(* IEC 61131-3 sources: stdmachine/plc/src/05_Sequencers, 11 files *)

(* ---- GVL_Active.st ---- *)
// Zone active du déploiement (docs/05 § 9 et § 10) : persistante, le PLC redémarre Stopped avec le dernier
// déploiement. À vérifier sur la cible : la taille (environ 1,5 Mo) des données persistantes.
{attribute 'qualified_only'}
VAR_GLOBAL PERSISTENT
    stMachine : ST_MachineData;
    aStation : ARRAY[1..GVL_Const.MAX_STATIONS] OF ST_StationData;
    aPressRecipe : ARRAY[1..GVL_Const.MAX_PRESS_RECIPES] OF ST_PressRecipe;
    bDeployed : BOOL;               // un déploiement a été activé
    nRetainId : ULINT;              // identifiant de la mémoire rémanente (docs/02 § 7.4), tiré au premier démarrage
END_VAR

(* ---- FB_GeneralSequencer.st ---- *)
// Séquenceur général (docs/05 § 5) : exécution du process général par mover, routage vers les stations des
// fonctions, files et priorités, préparation, fin d'opération (création et clôture des pièces, traces, qualité),
// table d'OF, fin des pièces en cours, variables de mover, mover à vider, mover hors service.
FUNCTION_BLOCK FB_GeneralSequencer
VAR_INPUT
    bDrain : BOOL;                  // fin des pièces en cours (docs/05 § 5.7), posé et levé par FB_Machine
END_VAR
VAR_OUTPUT
    bStopRequest : BOOL;            // impulsion : arrêt automatique demandé à la machine
    nStopReason : UINT;             // 1 OF terminé, 2 machine vidée, 3 arrêt qualité
    bMachineFault : BOOL;           // mover en défaut, alarme de process « défaut machine »
    nFaultCode : UINT;
END_VAR
VAR
    _refMachine : REFERENCE TO ST_MachineData;
    _refMgr : REFERENCE TO FB_MoverManager;
    _refQuality : REFERENCE TO FB_QualityMonitor;
    _refAlarms : REFERENCE TO FB_AlarmManager;
    _refTraces : REFERENCE TO FB_TraceBuffer;
    aStation : ARRAY[1..GVL_Const.MAX_STATIONS] OF POINTER TO FB_Station;
    _aLastReceived : ARRAY[1..GVL_Const.MAX_STATIONS] OF LINT;
    _aNoStationMs : ARRAY[1..GVL_Const.MAX_MOVERS] OF LREAL;
    _bExecute : BOOL;
    _bOrderDonePending : BOOL;      // l'OF actif vient de passer Done : arrêt quand plus aucune pièce
    _aGroupUsed : ARRAY[1..GVL_Const.MAX_GROUPS] OF BOOL;     // fonctions visées par une Route du process général
END_VAR
VAR PERSISTENT
    aMover : ARRAY[1..GVL_Const.MAX_MOVERS] OF ST_MoverCtx;
    aOrder : ARRAY[1..GVL_Const.MAX_ORDERS] OF ST_OrderState;
    nActiveOrder : USINT;           // rang dans aOrder, 0 = aucun
    _nReqSeq : UDINT;
    _nPartCounter : UDINT;
END_VAR

// ================================================================== mise en place

METHOD Init
VAR_INPUT
    refMachine : REFERENCE TO ST_MachineData;
    refMgr : REFERENCE TO FB_MoverManager;
    refQuality : REFERENCE TO FB_QualityMonitor;
    refAlarms : REFERENCE TO FB_AlarmManager;
    refTraces : REFERENCE TO FB_TraceBuffer;
END_VAR
_refMachine REF= refMachine;
_refMgr REF= refMgr;
_refQuality REF= refQuality;
_refAlarms REF= refAlarms;
_refTraces REF= refTraces;
END_METHOD

METHOD SetStation
VAR_INPUT
    nStation : USINT;
    pStation : POINTER TO FB_Station;
END_VAR
IF nStation >= 1 AND nStation <= GVL_Const.MAX_STATIONS THEN aStation[nStation] := pStation; END_IF
END_METHOD

// Reset machine (docs/05 § 6.3) : chaque mover détecté reçoit sa position ; les contextes et les pièces sont gardés
METHOD OnReset
VAR
    i : USINT;
    nPos : INT;
    ipDrv : I_PlanarDriver;
END_VAR
ipDrv := _refMgr.Driver;
FOR i := 1 TO _refMachine.nMovers DO
    aMover[i].bAbsent := FALSE;
    IF ipDrv <> 0 THEN
        IF NOT ipDrv.MoverDetected(i) THEN
            aMover[i].bAbsent := aMover[i].bOutOfService;       // D85 : un mover hors service peut être absent
            IF aMover[i].bAbsent AND __ISVALIDREF(_refAlarms) THEN _refAlarms.RaiseEvent(0, 915, i, E_Severity.Info); END_IF
        END_IF
    END_IF
    nPos := _refMgr.PositionAt(i);
    _refMgr.FreeAll(i, nPos);
    IF nPos > 0 THEN _refMgr.Reserve(nPos, i); END_IF
    aMover[i].nPos := nPos;
    CASE aMover[i].eState OF
        E_MoverState.Routing, E_MoverState.Halted, E_MoverState.Unknown, E_MoverState.Error:
            aMover[i].eState := E_MoverState.Ready;             // la Route en cours est reprise au Start
        E_MoverState.Queued:
            aMover[i].eState := E_MoverState.Buffered;
        E_MoverState.AtStation:
            IF NOT aMover[i].bStationAborted THEN
                aMover[i].eState := E_MoverState.Ready;
                aMover[i].bRequestPosted := FALSE;
            END_IF
    END_CASE
    IF aMover[i].nTable = 0 THEN
        aMover[i].nTable := 1;
        aMover[i].nPC := _refMachine.aTable[1].nStart;
    END_IF
END_FOR
END_METHOD

// Nouveau déploiement (docs/05 § 10) : variables de mover reprises par identifiant et type ; movers remis à
// l'étape 1 si le process général a changé de taille
METHOD OnDeploy
VAR_INPUT
    bRestartMovers : BOOL;
END_VAR
VAR
    i : USINT;
    v : USINT;
    k : USINT;
    stOld : ST_MoverCtx;
    bFound : BOOL;
END_VAR
FOR i := 1 TO GVL_Const.MAX_MOVERS DO
    stOld := aMover[i];
    FOR v := 1 TO GVL_Const.MAX_MOVER_VARS DO
        aMover[i].aVar[v] := 0;
        MEMSET(ADR(aMover[i].aVarPos[v]), 0, SIZEOF(ST_Position));
        aMover[i].aVarId[v] := 0;
        IF v <= _refMachine.nMoverVar THEN
            aMover[i].aVarId[v] := _refMachine.aMoverVar[v].nId;
            aMover[i].aVar[v] := _refMachine.aMoverVar[v].fInit;
            aMover[i].aVarPos[v] := _refMachine.aMoverVar[v].stInitPos;
            bFound := FALSE;
            IF _refMachine.aMoverVar[v].eReset <> E_MoverVarReset.OnDeploy THEN
                FOR k := 1 TO GVL_Const.MAX_MOVER_VARS DO
                    IF NOT bFound AND stOld.aVarId[k] = _refMachine.aMoverVar[v].nId AND stOld.aVarId[k] <> 0 THEN
                        aMover[i].aVar[v] := stOld.aVar[k];
                        aMover[i].aVarPos[v] := stOld.aVarPos[k];
                        bFound := TRUE;
                    END_IF
                END_FOR
            END_IF
        END_IF
    END_FOR
    IF bRestartMovers OR i > _refMachine.nMovers THEN
        aMover[i].nTable := 1;
        aMover[i].nPC := _refMachine.aTable[1].nStart;
        aMover[i].nDepth := 0;
        aMover[i].eState := E_MoverState.Ready;
        aMover[i].nTargetGroup := 0;
        aMover[i].bRequestPosted := FALSE;
    END_IF
END_FOR
IF bRestartMovers AND __ISVALIDREF(_refAlarms) THEN _refAlarms.RaiseEvent(0, 916, _refMachine.nMovers, E_Severity.Info); END_IF
ScanGroups();
END_METHOD

// ================================================================== cycle

METHOD Cycle
VAR_INPUT
    eState : E_State;               // état de la machine
END_VAR
VAR
    n : USINT;
    i : USINT;
    nArr : INT;
    nOldest : USINT;
END_VAR
_bExecute := eState = E_State.Execute;
bStopRequest := FALSE;
// Ordre des n°, en commençant par le mover qui attend depuis le plus longtemps (pas de famine)
nOldest := 1;
FOR i := 1 TO _refMachine.nMovers DO
    IF (aMover[i].eState = E_MoverState.Buffered OR aMover[i].eState = E_MoverState.Queued)
       AND (NOT (aMover[nOldest].eState = E_MoverState.Buffered OR aMover[nOldest].eState = E_MoverState.Queued) OR aMover[i].tWaitStart < aMover[nOldest].tWaitStart) THEN
        nOldest := i;
    END_IF
END_FOR
FOR n := 1 TO _refMachine.nMovers DO
    i := ((nOldest - 1 + n - 1) MOD _refMachine.nMovers) + 1;
    // Arrivées et timeouts, dans tous les états
    nArr := _refMgr.Arrived(i);
    IF nArr > 0 THEN _Arrive(i, nArr); END_IF
    IF _refMgr.TimedOut(i) AND aMover[i].eState <> E_MoverState.Error THEN
        aMover[i].eState := E_MoverState.Error;
        bMachineFault := TRUE;
        nFaultCode := 914;
        IF __ISVALIDREF(_refAlarms) THEN _refAlarms.RaiseEvent(0, 914, i, E_Severity.MachineFault); END_IF
    END_IF
    // Réaction qualité « mover hors service » (docs/10 § 5.1)
    aMover[i].bQualityLock := _refQuality.aMoverOut[i];

    IF _bExecute THEN
        IF (aMover[i].bOutOfService OR aMover[i].bQualityLock) AND aMover[i].eState = E_MoverState.Ready AND _Empty(i) THEN
            _SendToPark(i, FALSE);
        ELSIF aMover[i].bOutOfService AND aMover[i].bImmediate AND aMover[i].eState = E_MoverState.Ready AND NOT _Empty(i) THEN
            _SendToPark(i, TRUE);
        END_IF
        CASE aMover[i].eState OF
            E_MoverState.Ready: _RunMover(i);
            E_MoverState.Buffered:
                IF aMover[i].nTargetGroup = 0 THEN aMover[i].eState := E_MoverState.Ready; ELSE _TryRoute(i); END_IF
            E_MoverState.Queued: _Queued(i);
            E_MoverState.AtStation: _AtStation(i);
            E_MoverState.Halted: _Resume(i);
            E_MoverState.OutOfService:
                IF NOT aMover[i].bOutOfService AND NOT aMover[i].bQualityLock THEN _Restart(i); END_IF
        END_CASE
    ELSE
        // Held, Stopping : plus de nouveau routage ; les opérations lancées se terminent (docs/05 § 5.3)
        IF aMover[i].eState = E_MoverState.AtStation THEN _AtStation(i);
        ELSIF aMover[i].eState = E_MoverState.Ready OR aMover[i].eState = E_MoverState.Buffered OR aMover[i].eState = E_MoverState.Queued THEN
            IF eState = E_State.Held OR eState = E_State.Stopping THEN aMover[i].eWait := E_WaitReason.Held; END_IF
        END_IF
    END_IF
END_FOR
_CheckOrders();
IF bDrain AND (_bExecute OR eState = E_State.Held) AND PartsInProcess() = 0 AND NOT EntryInProgress() THEN
    bStopRequest := TRUE;
    nStopReason := 2;                                   // machine vidée (docs/05 § 5.7)
END_IF
IF _refQuality.bMachineStop THEN
    bStopRequest := TRUE;
    nStopReason := 3;
END_IF
_Publish();
END_METHOD

// ================================================================== process général d'un mover (docs/05 § 5.3)

METHOD PRIVATE _RunMover
VAR_INPUT
    i : USINT;
END_VAR
VAR
    m : REFERENCE TO ST_MoverCtx;
    ins : REFERENCE TO ST_Instr;
    nGuard : INT;
    n : INT;
    eSev : E_Severity;
END_VAR
m REF= aMover[i];
FOR nGuard := 1 TO 64 DO
    IF m.nPC < 1 OR m.nPC > _refMachine.nInstrCount THEN
        m.nTable := 1;
        m.nPC := _refMachine.aTable[1].nStart;
        RETURN;
    END_IF
    ins REF= _refMachine.aInstr[m.nPC];
    CASE ins.eOp OF
        E_Op.Jump:
            m.nPC := DINT_TO_INT(ins.aArg[1]);
        E_Op.JumpIfFalse:
            _MarkVerdictTested(i, DINT_TO_INT(ins.aArg[1]));
            IF _EvalCond(i, DINT_TO_INT(ins.aArg[1])) THEN m.nPC := m.nPC + 1; ELSE m.nPC := DINT_TO_INT(ins.aArg[2]); END_IF
        E_Op.SetVar:
            _SetVar(i);
            m.nPC := m.nPC + 1;
        E_Op.ResetMoverVars:
            _ResetVars(i, DINT_TO_INT(ins.aArg[1]));
            m.nPC := m.nPC + 1;
        E_Op.LoopInit:
            n := LIMIT(1, DINT_TO_INT(ins.aArg[1]), 8);
            m.aHidden[n] := _Resolve(i, ins.aParam[1]);
            m.nPC := m.nPC + 1;
        E_Op.LoopNext:
            n := LIMIT(1, DINT_TO_INT(ins.aArg[1]), 8);
            m.aHidden[n] := m.aHidden[n] - 1;
            IF m.aHidden[n] > 0 THEN m.nPC := DINT_TO_INT(ins.aArg[2]); ELSE m.nPC := m.nPC + 1; END_IF
        E_Op.Call:
            IF m.nDepth >= GVL_Const.MAX_CALL_DEPTH THEN
                m.eState := E_MoverState.Error;
                bMachineFault := TRUE;
                nFaultCode := 904;
                IF __ISVALIDREF(_refAlarms) THEN _refAlarms.RaiseEvent(0, 904, i, E_Severity.MachineFault); END_IF
                RETURN;
            END_IF
            m.nDepth := m.nDepth + 1;
            m.aRetTable[m.nDepth] := m.nTable;
            m.aRetPC[m.nDepth] := m.nPC + 1;
            m.nTable := DINT_TO_INT(ins.aArg[1]);
            m.nPC := _refMachine.aTable[m.nTable].nStart;
        E_Op.Return:
            IF m.nDepth = 0 THEN
                m.nTable := 1;
                m.nPC := _refMachine.aTable[1].nStart;
                RETURN;
            END_IF
            m.nTable := m.aRetTable[m.nDepth];
            m.nPC := m.aRetPC[m.nDepth];
            m.nDepth := m.nDepth - 1;
        E_Op.Alarm:
            // aArg[2] : 1 avertissement, sinon défaut machine (pas de station au niveau machine)
            IF ins.aArg[2] = 1 THEN eSev := E_Severity.Warning; ELSE eSev := E_Severity.MachineFault; END_IF
            IF __ISVALIDREF(_refAlarms) THEN _refAlarms.RaiseEvent(0, DINT_TO_UINT(ins.aArg[3]), i, eSev); END_IF
            IF ins.aArg[2] >= 2 THEN
                m.eState := E_MoverState.Error;
                bMachineFault := TRUE;
                nFaultCode := DINT_TO_UINT(ins.aArg[3]);
                RETURN;
            END_IF
            m.nPC := m.nPC + 1;
        E_Op.WaitCond:
            IF NOT _EvalCond(i, DINT_TO_INT(ins.aArg[1])) THEN RETURN; END_IF
            m.nPC := m.nPC + 1;
        E_Op.End:
            IF NOT _Empty(i) AND __ISVALIDREF(_refAlarms) THEN _refAlarms.RaiseEvent(0, 910, i, E_Severity.Warning); END_IF
            m.nTable := 1;
            m.nDepth := 0;
            m.nPC := _refMachine.aTable[1].nStart;
            RETURN;                                     // un tour de process par cycle au plus
        E_Op.Route:
            _StartRoute(i);
            RETURN;
    ELSE
        m.nPC := m.nPC + 1;                             // Nop, StepBegin, StepEnd
    END_CASE
END_FOR
END_METHOD

// ================================================================== routage (docs/05 § 5.4)

METHOD PRIVATE _StartRoute
VAR_INPUT
    i : USINT;
END_VAR
VAR
    m : REFERENCE TO ST_MoverCtx;
    ins : REFERENCE TO ST_Instr;
    nGroup : USINT;
    k : USINT;
    s : USINT;
    bBad : BOOL;
    bHandled : BOOL;
END_VAR
m REF= aMover[i];
ins REF= _refMachine.aInstr[m.nPC];
nGroup := DINT_TO_USINT(ins.aArg[1]);
m.nTargetOp := DINT_TO_USINT(ins.aArg[2]);
m.nTargetSlot := DINT_TO_USINT(ins.aArg[3]);
// 1. Pièce mauvaise non traitée par le process : redirection vers la fonction de rebut
FOR s := 1 TO GVL_Const.MAX_SLOTS DO
    IF m.aSlot[s].bPresent THEN
        bBad := bBad OR m.aSlot[s].aData[1] = 2;
        bHandled := bHandled OR m.aSlot[s].bBadHandled;
    END_IF
END_FOR
IF _refMachine.nRejectGroup > 0 AND nGroup <> _refMachine.nRejectGroup AND bBad AND NOT bHandled
   AND nGroup >= 1 AND nGroup <= GVL_Const.MAX_GROUPS AND_THEN _refMachine.aGroup[nGroup].eRole <> E_GroupRole.Reject THEN
    nGroup := _refMachine.nRejectGroup;
    m.nTargetOp := 1;
    MEMSET(ADR(m.aOpParam), 0, SIZEOF(m.aOpParam));
ELSE
    FOR k := 1 TO GVL_Const.MAX_PARAMS DO m.aOpParam[k] := _Resolve(i, ins.aParam[k]); END_FOR
END_IF
m.nTargetGroup := nGroup;
m.nStation := 0;
_aNoStationMs[i] := 0;
_TryRoute(i);
END_METHOD

METHOD PRIVATE _TryRoute
VAR_INPUT
    i : USINT;
END_VAR
VAR
    m : REFERENCE TO ST_MoverCtx;
    g : REFERENCE TO ST_GroupCfg;
    s : USINT;
    nBest : USINT;
    nLoad : INT;
    nBestLoad : INT;
    nDest : INT;
    k : USINT;
    eWait : E_WaitReason;
END_VAR
m REF= aMover[i];
IF m.nTargetGroup < 1 OR m.nTargetGroup > GVL_Const.MAX_GROUPS THEN m.eState := E_MoverState.Ready; RETURN; END_IF
g REF= _refMachine.aGroup[m.nTargetGroup];
// Fonction d'entrée : pas de chargement sans OF actif, OF complet, arrêt qualité du chargement, fin des pièces
IF g.eRole = E_GroupRole.Entry THEN
    eWait := _LoadingLock();
    IF eWait <> E_WaitReason.None THEN _WaitInBuffer(i, eWait); RETURN; END_IF
END_IF
// Candidates : stations membres en Execute, sans défaut, sans arrêt qualité, en production
nBest := 0;
IF NOT m.bOutOfService AND NOT m.bQualityLock THEN
    FOR s := 1 TO GVL_Const.MAX_STATIONS DO
        IF (SHR(g.nStationMask, s - 1) AND 1) = 1 AND_THEN _Routable(s) THEN
            nLoad := _LoadOf(s);
            IF nBest = 0 OR nLoad < nBestLoad OR (nLoad = nBestLoad AND _aLastReceived[s] < _aLastReceived[nBest]) THEN
                nBest := s;
                nBestLoad := nLoad;
            END_IF
        END_IF
    END_FOR
END_IF
IF nBest = 0 THEN
    _aNoStationMs[i] := _aNoStationMs[i] + F_CycleMs();
    IF (g.eRole = E_GroupRole.Reject OR _refMachine.nRejectGroup = 0) AND _aNoStationMs[i] > UDINT_TO_LREAL(_refMachine.nNoStationMs) AND NOT _Empty(i) THEN
        _SendToPark(i, TRUE);                       // mover à vider (911)
        RETURN;
    END_IF
    _WaitInBuffer(i, E_WaitReason.NoStation);
    RETURN;
END_IF
_aNoStationMs[i] := 0;
// Destination : position de travail libre et sans file, sinon une place de file, sinon un tampon
nDest := 0;
// (une position déjà tenue par ce mover compte comme libre : reprise après Reset)
IF _refMachine.aStation[nBest].nWorkPos > 0 AND_THEN _FreeFor(_refMachine.aStation[nBest].nWorkPos, i) AND NOT _HasQueue(nBest) THEN
    nDest := _refMachine.aStation[nBest].nWorkPos;
ELSE
    FOR k := 1 TO GVL_Const.MAX_QUEUE DO
        IF nDest = 0 AND _refMachine.aStation[nBest].aQueuePos[k] > 0 AND_THEN _FreeFor(_refMachine.aStation[nBest].aQueuePos[k], i) THEN
            nDest := _refMachine.aStation[nBest].aQueuePos[k];
        END_IF
    END_FOR
END_IF
IF nDest = 0 THEN
    _WaitInBuffer(i, E_WaitReason.NoStation);
    RETURN;
END_IF
_aLastReceived[nBest] := F_NowUtc();
m.nStation := nBest;
m.eWait := E_WaitReason.None;
IF _refMgr.MoveTo(i, nDest) THEN
    m.nDest := nDest;
    m.nPos := 0;
    m.eState := E_MoverState.Routing;
    m.bRequestPosted := FALSE;
    // Préparation : la demande est posée dès la réservation de la position de travail (docs/05 § 4.1)
    IF nDest = _refMachine.aStation[nBest].nWorkPos THEN _PostIfPrepare(i); END_IF
END_IF
END_METHOD

METHOD PRIVATE _FreeFor : BOOL
VAR_INPUT
    nPos : INT;
    i : USINT;
END_VAR
_FreeFor := _refMgr.Owner(nPos) = 0 OR _refMgr.Owner(nPos) = i;
END_METHOD

METHOD PRIVATE _LoadingLock : E_WaitReason
_LoadingLock := E_WaitReason.None;
IF _refQuality.bLoadingLocked THEN _LoadingLock := E_WaitReason.QualityStop;
ELSIF bDrain THEN _LoadingLock := E_WaitReason.Drain;
ELSIF nActiveOrder = 0 THEN _LoadingLock := E_WaitReason.NoOrder;
ELSIF aOrder[nActiveOrder].nGood + aOrder[nActiveOrder].nInProcess >= aOrder[nActiveOrder].nQuantity THEN _LoadingLock := E_WaitReason.OrderComplete;
END_IF
END_METHOD

METHOD PRIVATE _Routable : BOOL
VAR_INPUT
    s : USINT;
END_VAR
IF aStation[s] = 0 THEN _Routable := FALSE; RETURN; END_IF
_Routable := aStation[s]^.State = E_State.Execute AND NOT aStation[s]^.OutOfProduction AND NOT aStation[s]^.QualityLock
             AND _refMachine.aStation[s].bUsed;
END_METHOD

METHOD PRIVATE _LoadOf : INT
VAR_INPUT
    s : USINT;
END_VAR
VAR
    i : USINT;
END_VAR
_LoadOf := 0;
FOR i := 1 TO _refMachine.nMovers DO
    IF aMover[i].nStation = s THEN _LoadOf := _LoadOf + 1; END_IF
END_FOR
END_METHOD

METHOD PRIVATE _HasQueue : BOOL
VAR_INPUT
    s : USINT;
END_VAR
VAR
    i : USINT;
END_VAR
_HasQueue := FALSE;
FOR i := 1 TO _refMachine.nMovers DO
    IF aMover[i].nStation = s AND aMover[i].eState = E_MoverState.Queued THEN _HasQueue := TRUE; END_IF
END_FOR
END_METHOD

METHOD PRIVATE _WaitInBuffer
VAR_INPUT
    i : USINT;
    eReason : E_WaitReason;
END_VAR
VAR
    m : REFERENCE TO ST_MoverCtx;
    nBuf : INT;
END_VAR
m REF= aMover[i];
IF m.eState <> E_MoverState.Buffered THEN m.tWaitStart := F_NowUtc(); END_IF
m.eWait := eReason;
m.nStation := 0;
// Déjà sur un tampon ou au parcage : il y reste
IF m.nPos > 0 AND_THEN (_refMachine.aPlanarPos[m.nPos].eKind = E_PlanarPosKind.Buffer OR _refMachine.aPlanarPos[m.nPos].eKind = E_PlanarPosKind.Park) THEN
    m.eState := E_MoverState.Buffered;
    RETURN;
END_IF
IF m.eState = E_MoverState.Routing THEN RETURN; END_IF
nBuf := _refMgr.NearestFree(i, E_PlanarPosKind.Buffer);
IF nBuf > 0 AND_THEN _refMgr.MoveTo(i, nBuf) THEN
    m.nDest := nBuf;
    m.nPos := 0;
    m.eState := E_MoverState.Routing;
ELSE
    m.eState := E_MoverState.Buffered;                      // aucun tampon libre : il reste où il est
END_IF
END_METHOD

METHOD PRIVATE _SendToPark
VAR_INPUT
    i : USINT;
    bToEmpty : BOOL;
END_VAR
VAR
    m : REFERENCE TO ST_MoverCtx;
    nPark : INT;
END_VAR
m REF= aMover[i];
m.nStation := 0;
m.bToEmptyPark := bToEmpty;
IF bToEmpty AND __ISVALIDREF(_refAlarms) THEN _refAlarms.Raise(0, 911, i, E_Severity.Warning); END_IF
nPark := _refMachine.nParkPos;
IF nPark = 0 OR m.nPos = nPark THEN
    m.eState := SEL(bToEmpty OR NOT _Empty(i), E_MoverState.OutOfService, E_MoverState.ToEmpty);
    RETURN;
END_IF
IF _refMgr.MoveTo(i, nPark) THEN
    m.nDest := nPark;
    m.nPos := 0;
    m.eState := E_MoverState.Routing;
END_IF
END_METHOD

METHOD PRIVATE _Arrive
VAR_INPUT
    i : USINT;
    nPos : INT;
END_VAR
VAR
    m : REFERENCE TO ST_MoverCtx;
END_VAR
m REF= aMover[i];
m.nPos := nPos;
m.nDest := 0;
CASE _refMachine.aPlanarPos[nPos].eKind OF
    E_PlanarPosKind.Work:
        m.eState := E_MoverState.AtStation;
        IF m.bRequestPosted AND m.nStation >= 1 AND_THEN aStation[m.nStation] <> 0 THEN aStation[m.nStation]^.MoverArrived(m.nReqId); END_IF
    E_PlanarPosKind.Queue:
        // En Held et Stopping, le mover arrivé passe Halted (docs/05 § 5.3)
        IF _bExecute THEN m.eState := E_MoverState.Queued; ELSE m.eState := E_MoverState.Halted; END_IF
    E_PlanarPosKind.Buffer:
        IF _bExecute THEN m.eState := E_MoverState.Buffered; ELSE m.eState := E_MoverState.Halted; END_IF
    E_PlanarPosKind.Park:
        IF m.bToEmptyPark OR NOT _Empty(i) THEN m.eState := E_MoverState.ToEmpty; ELSE m.eState := E_MoverState.OutOfService; END_IF
END_CASE
m.tWaitStart := F_NowUtc();
END_METHOD

// Retour en Execute d'un mover Halted : il reprend selon la position où il se trouve, sans perdre son PC
METHOD PRIVATE _Resume
VAR_INPUT
    i : USINT;
END_VAR
VAR
    m : REFERENCE TO ST_MoverCtx;
END_VAR
m REF= aMover[i];
m.eWait := E_WaitReason.None;
IF m.nPos < 1 OR m.nPos > _refMachine.nPlanarPos OR m.nTargetGroup = 0 THEN
    m.eState := E_MoverState.Ready;
    RETURN;
END_IF
CASE _refMachine.aPlanarPos[m.nPos].eKind OF
    E_PlanarPosKind.Queue:
        IF m.nStation > 0 THEN m.eState := E_MoverState.Queued; ELSE m.eState := E_MoverState.Buffered; END_IF
    E_PlanarPosKind.Work:
        m.eState := E_MoverState.AtStation;
ELSE
    m.eState := E_MoverState.Buffered;
END_CASE
END_METHOD

// File : servie par priorité de la fonction visée (la plus haute d'abord), puis ordre d'arrivée
METHOD PRIVATE _Queued
VAR_INPUT
    i : USINT;
END_VAR
VAR
    m : REFERENCE TO ST_MoverCtx;
    s : USINT;
    j : USINT;
    nFirst : USINT;
    nWork : INT;
END_VAR
m REF= aMover[i];
s := m.nStation;
IF s < 1 OR s > GVL_Const.MAX_STATIONS OR_ELSE NOT _Routable(s) THEN
    m.eState := E_MoverState.Ready;                 // la station n'est plus disponible : le mover est réaffecté
    m.nStation := 0;
    RETURN;
END_IF
nWork := _refMachine.aStation[s].nWorkPos;
IF _refMgr.Owner(nWork) <> 0 THEN RETURN; END_IF
nFirst := 0;
FOR j := 1 TO _refMachine.nMovers DO
    IF aMover[j].eState = E_MoverState.Queued AND aMover[j].nStation = s THEN
        IF nFirst = 0 THEN
            nFirst := j;
        ELSIF _refMachine.aGroup[aMover[j].nTargetGroup].nPriority > _refMachine.aGroup[aMover[nFirst].nTargetGroup].nPriority
           OR (_refMachine.aGroup[aMover[j].nTargetGroup].nPriority = _refMachine.aGroup[aMover[nFirst].nTargetGroup].nPriority
               AND aMover[j].tWaitStart < aMover[nFirst].tWaitStart) THEN
            nFirst := j;
        END_IF
    END_IF
END_FOR
IF nFirst <> i THEN RETURN; END_IF
IF _refMgr.MoveTo(i, nWork) THEN
    m.nDest := nWork;
    m.nPos := 0;
    m.eState := E_MoverState.Routing;
    m.bRequestPosted := FALSE;
    _PostIfPrepare(i);
END_IF
END_METHOD

// ================================================================== demande d'opération

METHOD PRIVATE _PostIfPrepare
VAR_INPUT
    i : USINT;
END_VAR
VAR
    s : USINT;
END_VAR
s := aMover[i].nStation;
IF s < 1 OR s > GVL_Const.MAX_STATIONS OR_ELSE aStation[s] = 0 THEN RETURN; END_IF
IF aStation[s]^.PrepareWanted(aMover[i].nTargetGroup, aMover[i].nTargetOp) THEN _PostRequest(i, FALSE); END_IF
END_METHOD

METHOD PRIVATE _PostRequest : BOOL
VAR_INPUT
    i : USINT;
    bAtStation : BOOL;
END_VAR
VAR
    m : REFERENCE TO ST_MoverCtx;
    stReq : ST_OpRequest;
    s : USINT;
    k : USINT;
END_VAR
m REF= aMover[i];
s := m.nStation;
_PostRequest := FALSE;
IF s < 1 OR s > GVL_Const.MAX_STATIONS OR_ELSE aStation[s] = 0 THEN RETURN; END_IF
IF aStation[s]^.Response.eStatus <> E_OpStatus.Idle THEN RETURN; END_IF
_nReqSeq := _nReqSeq + 1;
stReq.nReqId := _nReqSeq;
stReq.nGroup := m.nTargetGroup;
stReq.nOperation := m.nTargetOp;
stReq.nMover := i;
stReq.nSlot := m.nTargetSlot;
stReq.bMoverAtStation := bAtStation;
stReq.aParam := m.aOpParam;
IF aStation[s]^.Offer(stReq, ADR(aMover[i])) THEN
    m.nReqId := stReq.nReqId;
    m.bRequestPosted := TRUE;
    m.tOpStart := F_NowUtc();
    FOR k := 1 TO GVL_Const.MAX_SLOTS DO
        m.aBadAtArrival[k] := m.aSlot[k].bPresent AND m.aSlot[k].aData[1] = 2;
    END_FOR
    _PostRequest := TRUE;
END_IF
END_METHOD

METHOD PRIVATE _AtStation
VAR_INPUT
    i : USINT;
END_VAR
VAR
    m : REFERENCE TO ST_MoverCtx;
    s : USINT;
    k : USINT;
    eSt : E_State;
END_VAR
m REF= aMover[i];
s := m.nStation;
IF s < 1 OR s > GVL_Const.MAX_STATIONS OR_ELSE aStation[s] = 0 THEN m.eState := E_MoverState.Ready; RETURN; END_IF
eSt := aStation[s]^.State;
IF m.bStationAborted THEN
    // Le mover reste en position de travail jusqu'à la fin du Clearing, puis part au rebut (docs/05 § 6.4)
    IF eSt = E_State.Stopped OR eSt = E_State.Idle OR eSt = E_State.Execute THEN
        m.bStationAborted := FALSE;
        m.bRequestPosted := FALSE;
        m.nStation := 0;
        m.eState := E_MoverState.Ready;
    END_IF
    RETURN;
END_IF
IF NOT m.bRequestPosted THEN
    IF _bExecute AND eSt = E_State.Execute AND _Routable(s) THEN _PostRequest(i, TRUE); END_IF
    RETURN;
END_IF
IF aStation[s]^.Response.nReqId <> m.nReqId THEN RETURN; END_IF
CASE aStation[s]^.Response.eStatus OF
    E_OpStatus.Done, E_OpStatus.Failed:
        _FinishOperation(i);
    E_OpStatus.Aborted:
        IF aStation[s]^.Response.nErrorCode = 907 THEN
            // Préparation annulée par l'arrêt : rien n'a touché la pièce, le mover reprend sa Route au Start suivant
            m.bRequestPosted := FALSE;
            m.nStation := 0;
            m.eState := E_MoverState.Ready;
        ELSE
            // Station Aborted : pièces mauvaises, la position de travail reste tenue (docs/05 § 6.4)
            FOR k := 1 TO GVL_Const.MAX_SLOTS DO
                IF m.aSlot[k].bPresent THEN
                    m.aSlot[k].aData[1] := 2;
                    m.aSlot[k].bBadHandled := FALSE;
                    m.aDefectBad[k] := TRUE;
                END_IF
            END_FOR
            m.bStationAborted := TRUE;
        END_IF
        aStation[s]^.AckResponse();
END_CASE
END_METHOD

// ================================================================== fin d'une opération (docs/05 § 5.5)

METHOD PRIVATE _FinishOperation
VAR_INPUT
    i : USINT;
END_VAR
VAR
    m : REFERENCE TO ST_MoverCtx;
    g : REFERENCE TO ST_GroupCfg;
    ins : REFERENCE TO ST_Instr;
    st : POINTER TO FB_Station;
    s : USINT;
    k : USINT;
    j : USINT;
    bFailed : BOOL;
    bBad : BOOL;
    bClosed : BOOL;
    bClosedBad : BOOL;
    nFirst : USINT;
    nLast : USINT;
    nImpute : UINT;
    nOrderIdx : USINT;
    stTrace : ST_TraceRecord;
END_VAR
m REF= aMover[i];
s := m.nStation;
st := aStation[s];
g REF= _refMachine.aGroup[m.nTargetGroup];
ins REF= _refMachine.aInstr[m.nPC];
bFailed := st^.Response.eStatus = E_OpStatus.Failed;

// 0. Sorties de l'opération vers les cibles de la Route (docs/02 § 5.5)
IF NOT bFailed THEN
    FOR k := 1 TO GVL_Const.MAX_OUTPUTS DO
        IF (SHR(st^.Response.nOutMask, k - 1) AND 1) = 1 THEN _BindOutput(i, ins.aBind[k], st^.Response.aOut[k], st^.Response.stOutPos); END_IF
    END_FOR
END_IF
st^.AckResponse();

// 1. Libérer la position de travail (la file est promue par _Queued)
_refMgr.Free(m.nPos, i);
m.nPos := 0;
m.nStation := 0;
m.bRequestPosted := FALSE;

IF m.nTargetSlot = 0 THEN nFirst := 1; nLast := _refMachine.nSlots; ELSE nFirst := m.nTargetSlot; nLast := m.nTargetSlot; END_IF
FOR k := nFirst TO MIN(nLast, GVL_Const.MAX_SLOTS) DO
    // 2. Création des pièces par une opération d'entrée réussie
    IF g.eRole = E_GroupRole.Entry AND NOT bFailed AND NOT m.aSlot[k].bPresent AND nActiveOrder > 0 THEN
        m.aSlot[k].bPresent := TRUE;
        _nPartCounter := _nPartCounter + 1;
        IF LEN(m.aSlot[k].sPartId) = 0 THEN m.aSlot[k].sPartId := F_PartId(_refMachine.sMachineName, _nPartCounter); END_IF
        m.aSlot[k].eStatus := E_PartStatus.InProcess;
        m.aSlot[k].nOrder := aOrder[nActiveOrder].nOrder;
        m.aSlot[k].tCreated := F_NowUtc();
        m.aSlot[k].nOps := 0;
        m.aSlot[k].bBadHandled := FALSE;
        aOrder[nActiveOrder].nInProcess := aOrder[nActiveOrder].nInProcess + 1;
        m.aBadAtArrival[k] := FALSE;
        m.aDefectBad[k] := FALSE;
    END_IF
    IF m.aSlot[k].bPresent THEN
        IF bFailed THEN m.aSlot[k].aData[1] := 2; END_IF
        bBad := m.aSlot[k].aData[1] = 2;
        IF m.aSlot[k].nOps < GVL_Const.MAX_PART_OPS THEN
            m.aSlot[k].nOps := m.aSlot[k].nOps + 1;
            m.aSlot[k].aOps[m.aSlot[k].nOps].nStation := s;
            m.aSlot[k].aOps[m.aSlot[k].nOps].nGroup := m.nTargetGroup;
            m.aSlot[k].aOps[m.aSlot[k].nOps].eVerdictAfter := F_Verdict(m.aSlot[k].aData[1]);
        END_IF
        // 6. Surveillance des rebuts : un verdict déjà mauvais à l'arrivée ne compte pas pour cette station
        IF NOT m.aBadAtArrival[k] AND NOT m.aDefectBad[k] THEN
            _refQuality.Record(E_QualityScope.Station, s, bBad);
            _refQuality.Record(E_QualityScope.Group, m.nTargetGroup, bBad);
            nImpute := _refMachine.stQuality.aGroupImpute[m.nTargetGroup];
            IF nImpute <> 0 THEN
                FOR j := 1 TO m.aSlot[k].nOps - 1 DO
                    IF (SHR(nImpute, m.aSlot[k].aOps[j].nGroup - 1) AND 1) = 1 THEN
                        _refQuality.Record(E_QualityScope.StationImputed, m.aSlot[k].aOps[j].nStation, bBad);
                    END_IF
                END_FOR
            END_IF
        END_IF
        // 3 et 4. Clôture : pièce retirée par l'opération, sortie, rebut
        bClosed := FALSE;
        bClosedBad := FALSE;
        IF m.aSlot[k].eStatus = E_PartStatus.Removed THEN
            bClosed := TRUE;
            bClosedBad := TRUE;
        ELSIF g.eRole = E_GroupRole.Exit AND NOT bFailed THEN
            bClosed := TRUE;
            m.aSlot[k].eStatus := E_PartStatus.Exited;
        ELSIF g.eRole = E_GroupRole.Reject THEN
            bClosed := TRUE;
            bClosedBad := TRUE;
            m.aSlot[k].eStatus := E_PartStatus.Rejected;
        END_IF
        IF bClosed AND NOT m.aDefectBad[k] THEN
            _refQuality.Record(E_QualityScope.Mover, i, bClosedBad OR bBad);
            _refQuality.Record(E_QualityScope.Machine, 0, bClosedBad OR bBad);
        END_IF
        // 5. Trace
        MEMSET(ADR(stTrace), 0, SIZEOF(stTrace));
        stTrace.sPartId := m.aSlot[k].sPartId;
        stTrace.nOrder := m.aSlot[k].nOrder;
        stTrace.nMover := i;
        stTrace.nSlot := k;
        stTrace.nStation := s;
        stTrace.nGroup := m.nTargetGroup;
        stTrace.nOperation := m.nTargetOp;
        stTrace.tStart := m.tOpStart;
        stTrace.tEnd := F_NowUtc();
        stTrace.eVerdict := F_Verdict(m.aSlot[k].aData[1]);
        stTrace.nErrorCode := st^.Response.nErrorCode;
        stTrace.aData := m.aSlot[k].aData;
        // Courbe de presse enregistrée par la station pendant cette opération (docs/05 § 9)
        IF GVL_Curves.aLastCurveId[s] <> 0 AND GVL_Curves.aLastCurveTime[s] >= m.tOpStart THEN stTrace.nCurveId := GVL_Curves.aLastCurveId[s]; END_IF
        _refTraces.Add(stTrace);
        IF bClosed THEN
            nOrderIdx := _OrderIndex(m.aSlot[k].nOrder);
            IF nOrderIdx > 0 THEN _CloseOrderPart(nOrderIdx, bClosedBad OR bBad); END_IF
            MEMSET(ADR(m.aSlot[k]), 0, SIZEOF(m.aSlot[k]));
            m.aDefectBad[k] := FALSE;
            m.aBadAtArrival[k] := FALSE;
        END_IF
    END_IF
END_FOR
IF _Empty(i) THEN _ResetOnEmpty(i); END_IF

// 7. Avancer le PC ; le parcage d'un mover verrouillé et vide est traité au cycle suivant
m.nPC := m.nPC + 1;
m.eState := E_MoverState.Ready;
m.nTargetGroup := 0;
END_METHOD

METHOD PRIVATE _BindOutput
VAR_INPUT
    i : USINT;
    stBind : ST_Bind;
    fValue : LREAL;
    stPos : ST_Position;
END_VAR
VAR
    n : INT;
    k : USINT;
END_VAR
n := stBind.nIndex;
CASE stBind.eTarget OF
    E_BindTarget.PartData:
        FOR k := 1 TO GVL_Const.MAX_SLOTS DO
            IF aMover[i].aSlot[k].bPresent AND n >= 1 AND n <= GVL_Const.MAX_PART_DATA AND (aMover[i].nTargetSlot = 0 OR aMover[i].nTargetSlot = k) THEN
                aMover[i].aSlot[k].aData[n] := fValue;
            END_IF
        END_FOR
    E_BindTarget.Verdict:
        FOR k := 1 TO GVL_Const.MAX_SLOTS DO
            IF aMover[i].aSlot[k].bPresent AND (aMover[i].nTargetSlot = 0 OR aMover[i].nTargetSlot = k) THEN aMover[i].aSlot[k].aData[1] := fValue; END_IF
        END_FOR
    E_BindTarget.MoverData:
        IF n >= 1 AND n <= _refMachine.nMoverVar THEN
            IF _refMachine.aMoverVar[n].eType = E_VarType.Position THEN aMover[i].aVarPos[n] := stPos; ELSE aMover[i].aVar[n] := fValue; END_IF
        END_IF
END_CASE
END_METHOD

// Variables de mover à règle « quand le mover est vide » (docs/05 § 5.8)
METHOD PRIVATE _ResetOnEmpty
VAR_INPUT
    i : USINT;
END_VAR
VAR
    v : USINT;
END_VAR
FOR v := 1 TO _refMachine.nMoverVar DO
    IF _refMachine.aMoverVar[v].eReset = E_MoverVarReset.OnEmpty THEN
        aMover[i].aVar[v] := _refMachine.aMoverVar[v].fInit;
        aMover[i].aVarPos[v] := _refMachine.aMoverVar[v].stInitPos;
    END_IF
END_FOR
END_METHOD

METHOD PRIVATE _ResetVars
VAR_INPUT
    i : USINT;
    nRank : INT;
END_VAR
VAR
    v : INT;
END_VAR
FOR v := 1 TO _refMachine.nMoverVar DO
    IF (nRank = 0 AND _refMachine.aMoverVar[v].eReset <> E_MoverVarReset.Never) OR nRank = v THEN
        aMover[i].aVar[v] := _refMachine.aMoverVar[v].fInit;
        aMover[i].aVarPos[v] := _refMachine.aMoverVar[v].stInitPos;
    END_IF
END_FOR
END_METHOD

METHOD PRIVATE _Restart
VAR_INPUT
    i : USINT;
END_VAR
aMover[i].nTable := 1;
aMover[i].nDepth := 0;
aMover[i].nPC := _refMachine.aTable[1].nStart;
aMover[i].nTargetGroup := 0;
aMover[i].eState := E_MoverState.Ready;
aMover[i].eWait := E_WaitReason.None;
aMover[i].bToEmptyPark := FALSE;
END_METHOD

// ================================================================== valeurs et conditions du process général

METHOD PRIVATE _FirstPart : POINTER TO ST_Part
VAR_INPUT
    i : USINT;
END_VAR
VAR
    k : USINT;
END_VAR
_FirstPart := ADR(aMover[i].aSlot[1]);
FOR k := 1 TO GVL_Const.MAX_SLOTS DO
    IF aMover[i].aSlot[k].bPresent THEN _FirstPart := ADR(aMover[i].aSlot[k]); RETURN; END_IF
END_FOR
END_METHOD

METHOD PRIVATE _Resolve : LREAL
VAR_INPUT
    i : USINT;
    stVal : ST_Value;
END_VAR
VAR
    pPart : POINTER TO ST_Part;
    n : INT;
    nIdx : USINT;
END_VAR
n := stVal.nIndex;
CASE stVal.eSource OF
    E_ValueSource.Const:
        _Resolve := stVal.fValue;
    E_ValueSource.PartData:
        pPart := _FirstPart(i);
        IF n >= 1 AND n <= GVL_Const.MAX_PART_DATA THEN _Resolve := pPart^.aData[n]; END_IF
    E_ValueSource.MoverData:
        IF n >= 1 AND n <= GVL_Const.MAX_MOVER_VARS THEN _Resolve := aMover[i].aVar[n]; END_IF
    E_ValueSource.OrderParam:
        // OF de la première pièce présente, sinon l'OF actif (opération d'entrée) (docs/05 § 5.6)
        pPart := _FirstPart(i);
        nIdx := 0;
        IF pPart^.bPresent THEN nIdx := _OrderIndex(pPart^.nOrder); END_IF
        IF nIdx = 0 THEN nIdx := nActiveOrder; END_IF
        IF nIdx > 0 AND n >= 1 AND n <= GVL_Const.MAX_ORDER_PARAMS THEN _Resolve := aOrder[nIdx].aParam[n]; END_IF
    E_ValueSource.System:
        CASE n OF
            1: _Resolve := 1.0;                                     // mover présent
            3:
                pPart := _FirstPart(i);
                IF pPart^.bPresent THEN _Resolve := UDINT_TO_LREAL(pPart^.nOrder); END_IF
        END_CASE
    E_ValueSource.Speed:
        _Resolve := INT_TO_LREAL(n);
END_CASE
END_METHOD

METHOD PRIVATE _EvalCond : BOOL
VAR_INPUT
    i : USINT;
    n : INT;
END_VAR
VAR
    k : USINT;
    r : BOOL;
    bAll : BOOL;
END_VAR
IF n < 1 OR n > GVL_Const.MAX_COND THEN _EvalCond := TRUE; RETURN; END_IF
IF _refMachine.aCond[n].nTerms = 0 THEN _EvalCond := TRUE; RETURN; END_IF
bAll := _refMachine.aCond[n].eCombine = E_Combine.All;
FOR k := 1 TO MIN(_refMachine.aCond[n].nTerms, GVL_Const.MAX_COND_TERMS) DO
    r := F_Compare(_Resolve(i, _refMachine.aCond[n].aTerm[k].stLeft), _refMachine.aCond[n].aTerm[k].eCmp, _Resolve(i, _refMachine.aCond[n].aTerm[k].stRight));
    IF bAll AND NOT r THEN _EvalCond := FALSE; RETURN; END_IF
    IF NOT bAll AND r THEN _EvalCond := TRUE; RETURN; END_IF
END_FOR
_EvalCond := bAll;
END_METHOD

// Un Si qui teste le verdict traite lui-même la pièce mauvaise : pas de redirection automatique (docs/02 § 6.2)
METHOD PRIVATE _MarkVerdictTested
VAR_INPUT
    i : USINT;
    n : INT;
END_VAR
VAR
    k : USINT;
    s : USINT;
    bTested : BOOL;
END_VAR
IF n < 1 OR n > GVL_Const.MAX_COND THEN RETURN; END_IF
FOR k := 1 TO MIN(_refMachine.aCond[n].nTerms, GVL_Const.MAX_COND_TERMS) DO
    bTested := bTested
        OR (_refMachine.aCond[n].aTerm[k].stLeft.eSource = E_ValueSource.PartData AND _refMachine.aCond[n].aTerm[k].stLeft.nIndex = 1)
        OR (_refMachine.aCond[n].aTerm[k].stRight.eSource = E_ValueSource.PartData AND _refMachine.aCond[n].aTerm[k].stRight.nIndex = 1);
END_FOR
// Seul un test fait pendant que la pièce est mauvaise la traite (« depuis qu'il est devenu mauvais »)
IF bTested THEN
    FOR s := 1 TO GVL_Const.MAX_SLOTS DO
        IF aMover[i].aSlot[s].bPresent AND aMover[i].aSlot[s].aData[1] = 2 THEN aMover[i].aSlot[s].bBadHandled := TRUE; END_IF
    END_FOR
END_IF
END_METHOD

METHOD PRIVATE _SetVar
VAR_INPUT
    i : USINT;
END_VAR
VAR
    ins : REFERENCE TO ST_Instr;
    pPart : POINTER TO ST_Part;
    fValue : LREAL;
    n : INT;
END_VAR
ins REF= _refMachine.aInstr[aMover[i].nPC];
fValue := _Resolve(i, ins.aParam[1]);
n := ins.aBind[1].nIndex;
CASE ins.aBind[1].eTarget OF
    E_BindTarget.PartData:
        pPart := _FirstPart(i);
        IF pPart^.bPresent AND n >= 1 AND n <= GVL_Const.MAX_PART_DATA THEN pPart^.aData[n] := F_ApplyOp(pPart^.aData[n], fValue, ins.aArg[1]); END_IF
    E_BindTarget.Verdict:
        pPart := _FirstPart(i);
        IF pPart^.bPresent THEN pPart^.aData[1] := fValue; END_IF
    E_BindTarget.MoverData:
        IF n >= 1 AND n <= GVL_Const.MAX_MOVER_VARS THEN aMover[i].aVar[n] := F_ApplyOp(aMover[i].aVar[n], fValue, ins.aArg[1]); END_IF
END_CASE
END_METHOD

METHOD PRIVATE _Empty : BOOL
VAR_INPUT
    i : USINT;
END_VAR
VAR
    k : USINT;
END_VAR
_Empty := TRUE;
FOR k := 1 TO GVL_Const.MAX_SLOTS DO
    IF aMover[i].aSlot[k].bPresent THEN _Empty := FALSE; END_IF
END_FOR
END_METHOD

// ================================================================== OF (docs/05 § 5.6)

METHOD Activate : E_RejectReason
VAR_INPUT
    stReq : ST_OrderRequest;
END_VAR
VAR
    nIdx : USINT;
    k : USINT;
    bNewReference : BOOL;
END_VAR
nIdx := _OrderIndex(stReq.nOrder);
IF nIdx = 0 THEN
    FOR k := 1 TO GVL_Const.MAX_ORDERS DO
        // Place libre, ou OF terminé ou suspendu sans pièce en cours (il quitte la table, la HMI garde ses compteurs)
        IF nIdx = 0 AND k <> nActiveOrder AND (aOrder[k].eState = E_OrderState.Free
           OR ((aOrder[k].eState = E_OrderState.Done OR aOrder[k].eState = E_OrderState.Suspended) AND aOrder[k].nInProcess = 0)) THEN
            nIdx := k;
        END_IF
    END_FOR
    IF nIdx = 0 THEN Activate := E_RejectReason.TableFull; RETURN; END_IF
    MEMSET(ADR(aOrder[nIdx]), 0, SIZEOF(aOrder[nIdx]));
    aOrder[nIdx].nOrder := stReq.nOrder;
    aOrder[nIdx].nGood := stReq.nGoodDone;
    aOrder[nIdx].nBad := stReq.nBadDone;
END_IF
bNewReference := nActiveOrder = 0 OR_ELSE aOrder[nActiveOrder].sReference <> stReq.sReference;
IF nActiveOrder > 0 AND nActiveOrder <> nIdx AND aOrder[nActiveOrder].eState = E_OrderState.Active THEN
    aOrder[nActiveOrder].eState := E_OrderState.Suspended;
END_IF
aOrder[nIdx].sNumber := stReq.sNumber;
aOrder[nIdx].sReference := stReq.sReference;
aOrder[nIdx].nQuantity := stReq.nQuantity;
aOrder[nIdx].aParam := stReq.aParam;
aOrder[nIdx].eState := E_OrderState.Active;
nActiveOrder := nIdx;
_bOrderDonePending := FALSE;
IF bNewReference THEN _refQuality.ResetAllWindows(); END_IF      // D87
FOR k := 1 TO GVL_Const.MAX_STATIONS DO
    IF aStation[k] <> 0 THEN aStation[k]^.OnOrderChange(); END_IF
END_FOR
Activate := E_RejectReason.None;
END_METHOD

METHOD Suspend : E_RejectReason
IF nActiveOrder = 0 THEN Suspend := E_RejectReason.NotConfigured; RETURN; END_IF
IF aOrder[nActiveOrder].eState = E_OrderState.Active THEN aOrder[nActiveOrder].eState := E_OrderState.Suspended; END_IF
nActiveOrder := 0;
Suspend := E_RejectReason.None;
END_METHOD

METHOD Cancel : E_RejectReason
VAR_INPUT
    nOrder : UDINT;
END_VAR
VAR
    nIdx : USINT;
END_VAR
nIdx := _OrderIndex(nOrder);
IF nIdx = 0 THEN Cancel := E_RejectReason.NotConfigured; RETURN; END_IF
IF aOrder[nIdx].nInProcess > 0 THEN Cancel := E_RejectReason.PartsInProcess; RETURN; END_IF
IF nActiveOrder = nIdx THEN nActiveOrder := 0; END_IF
MEMSET(ADR(aOrder[nIdx]), 0, SIZEOF(aOrder[nIdx]));
Cancel := E_RejectReason.None;
END_METHOD

METHOD PRIVATE _OrderIndex : USINT
VAR_INPUT
    nOrder : UDINT;
END_VAR
VAR
    k : USINT;
END_VAR
_OrderIndex := 0;
IF nOrder = 0 THEN RETURN; END_IF
FOR k := 1 TO GVL_Const.MAX_ORDERS DO
    IF aOrder[k].nOrder = nOrder AND aOrder[k].eState <> E_OrderState.Free THEN _OrderIndex := k; RETURN; END_IF
END_FOR
END_METHOD

METHOD PRIVATE _CloseOrderPart
VAR_INPUT
    nIdx : USINT;
    bBad : BOOL;
END_VAR
IF aOrder[nIdx].nInProcess > 0 THEN aOrder[nIdx].nInProcess := aOrder[nIdx].nInProcess - 1; END_IF
IF bBad THEN aOrder[nIdx].nBad := aOrder[nIdx].nBad + 1; ELSE aOrder[nIdx].nGood := aOrder[nIdx].nGood + 1; END_IF
_refQuality.RecordOrder(aOrder[nIdx], bBad);
END_METHOD

METHOD PRIVATE _CheckOrders
VAR
    k : USINT;
END_VAR
// Un OF complet dont plus aucune pièce n'est en cours passe Done, actif ou suspendu (docs/05 § 5.6)
FOR k := 1 TO GVL_Const.MAX_ORDERS DO
    IF (aOrder[k].eState = E_OrderState.Active OR aOrder[k].eState = E_OrderState.Suspended)
       AND aOrder[k].nGood + aOrder[k].nInProcess >= aOrder[k].nQuantity AND aOrder[k].nInProcess = 0 THEN
        aOrder[k].eState := E_OrderState.Done;
        IF k = nActiveOrder THEN _bOrderDonePending := TRUE; END_IF
    END_IF
END_FOR
// OF actif terminé : arrêt automatique dès qu'aucune pièce d'aucun OF n'est en cours
IF _bOrderDonePending AND _bExecute AND PartsInProcess() = 0 THEN
    _bOrderDonePending := FALSE;
    bStopRequest := TRUE;
    nStopReason := 1;                               // événement « OF terminé » (raison d'arrêt)
END_IF
END_METHOD

// ================================================================== commandes HMI

// Retrait des pièces d'un mover à vider confirmé par l'opérateur (docs/02 § 10)
METHOD ConfirmRemoved : E_RejectReason
VAR_INPUT
    nMover : USINT;
END_VAR
VAR
    k : USINT;
    nIdx : USINT;
END_VAR
IF nMover < 1 OR nMover > _refMachine.nMovers THEN ConfirmRemoved := E_RejectReason.NotConfigured; RETURN; END_IF
IF aMover[nMover].eState <> E_MoverState.ToEmpty THEN ConfirmRemoved := E_RejectReason.WrongState; RETURN; END_IF
FOR k := 1 TO GVL_Const.MAX_SLOTS DO
    IF aMover[nMover].aSlot[k].bPresent THEN
        nIdx := _OrderIndex(aMover[nMover].aSlot[k].nOrder);
        IF nIdx > 0 THEN _CloseOrderPart(nIdx, TRUE); END_IF       // retrait manuel : compte dans le budget d'OF
        MEMSET(ADR(aMover[nMover].aSlot[k]), 0, SIZEOF(aMover[nMover].aSlot[k]));
    END_IF
END_FOR
_ResetOnEmpty(nMover);
IF aMover[nMover].bOutOfService OR aMover[nMover].bQualityLock THEN
    aMover[nMover].eState := E_MoverState.OutOfService;
ELSE
    _Restart(nMover);
END_IF
// Une seule alarme 911 pour la machine : elle tombe quand plus aucun mover n'est à vider
IF NOT AnyToEmpty() AND __ISVALIDREF(_refAlarms) THEN _refAlarms.Clear(0, 911); END_IF
ConfirmRemoved := E_RejectReason.None;
END_METHOD

METHOD SetMoverVar : E_RejectReason
VAR_INPUT
    stReq : ST_MoverVarRequest;
END_VAR
IF stReq.nMover < 1 OR stReq.nMover > _refMachine.nMovers OR stReq.nVar < 1 OR stReq.nVar > _refMachine.nMoverVar THEN
    SetMoverVar := E_RejectReason.NotConfigured;
    RETURN;
END_IF
IF stReq.bReset THEN
    aMover[stReq.nMover].aVar[stReq.nVar] := _refMachine.aMoverVar[stReq.nVar].fInit;
    aMover[stReq.nMover].aVarPos[stReq.nVar] := _refMachine.aMoverVar[stReq.nVar].stInitPos;
ELSIF _refMachine.aMoverVar[stReq.nVar].eType = E_VarType.Position THEN
    aMover[stReq.nMover].aVarPos[stReq.nVar] := stReq.stPos;
ELSE
    aMover[stReq.nMover].aVar[stReq.nVar] := stReq.fValue;
END_IF
SetMoverVar := E_RejectReason.None;
END_METHOD

METHOD SetOutOfService
VAR_INPUT
    nMover : USINT;
    bOut : BOOL;
    bImmediate : BOOL;
END_VAR
IF nMover < 1 OR nMover > GVL_Const.MAX_MOVERS THEN RETURN; END_IF
aMover[nMover].bOutOfService := bOut;
aMover[nMover].bImmediate := bOut AND bImmediate;
IF NOT bOut AND aMover[nMover].eState = E_MoverState.OutOfService AND NOT aMover[nMover].bQualityLock THEN _Restart(nMover); END_IF
END_METHOD

// ================================================================== état

METHOD PartsInProcess : UINT
VAR
    i : USINT;
    k : USINT;
END_VAR
PartsInProcess := 0;
FOR i := 1 TO _refMachine.nMovers DO
    FOR k := 1 TO GVL_Const.MAX_SLOTS DO
        IF aMover[i].aSlot[k].bPresent THEN PartsInProcess := PartsInProcess + 1; END_IF
    END_FOR
END_FOR
END_METHOD

// Une opération d'entrée est-elle en cours ou engagée ? (fin des pièces : on la laisse finir, docs/05 § 5.7)
METHOD EntryInProgress : BOOL
VAR
    i : USINT;
END_VAR
EntryInProgress := FALSE;
FOR i := 1 TO _refMachine.nMovers DO
    IF aMover[i].nTargetGroup >= 1 AND aMover[i].nTargetGroup <= GVL_Const.MAX_GROUPS THEN
        IF _refMachine.aGroup[aMover[i].nTargetGroup].eRole = E_GroupRole.Entry
           AND (aMover[i].bRequestPosted OR aMover[i].eState = E_MoverState.AtStation OR (aMover[i].eState = E_MoverState.Routing AND aMover[i].nStation > 0)) THEN
            EntryInProgress := TRUE;
        END_IF
    END_IF
END_FOR
END_METHOD

METHOD AnyAtStation : BOOL
VAR
    i : USINT;
END_VAR
AnyAtStation := FALSE;
FOR i := 1 TO _refMachine.nMovers DO
    IF aMover[i].eState = E_MoverState.AtStation AND aMover[i].bRequestPosted THEN AnyAtStation := TRUE; END_IF
END_FOR
END_METHOD

METHOD AnyToEmpty : BOOL
VAR
    i : USINT;
END_VAR
AnyToEmpty := FALSE;
FOR i := 1 TO _refMachine.nMovers DO
    IF aMover[i].eState = E_MoverState.ToEmpty THEN AnyToEmpty := TRUE; END_IF
END_FOR
END_METHOD

// Fonction utilisée par le process général à laquelle il manque une station (docs/05 § 5.2) ; 0 = aucune.
// nCheck 1 : aucune station disponible (pas Aborted ni Stopped), défaut 913 en Execute ;
// nCheck 2 : aucune station en Idle (Resetting → Idle) ; nCheck 3 : toutes ses stations Aborted (Resetting).
// Une station volontairement retirée (hors production, arrêt qualité) ne déclenche jamais le défaut.
METHOD MissingGroup : USINT
VAR_INPUT
    nCheck : USINT;
END_VAR
VAR
    g : USINT;
    s : USINT;
    bOk : BOOL;
    bAny : BOOL;
    bWithdrawn : BOOL;
    eSt : E_State;
END_VAR
MissingGroup := 0;
FOR g := 1 TO GVL_Const.MAX_GROUPS DO
    IF _aGroupUsed[g] THEN
        bOk := FALSE;
        bAny := FALSE;
        bWithdrawn := FALSE;
        FOR s := 1 TO GVL_Const.MAX_STATIONS DO
            IF (SHR(_refMachine.aGroup[g].nStationMask, s - 1) AND 1) = 1 AND_THEN aStation[s] <> 0 THEN
                bAny := TRUE;
                eSt := aStation[s]^.State;
                IF aStation[s]^.OutOfProduction OR aStation[s]^.QualityLock THEN
                    bWithdrawn := TRUE;
                END_IF
                CASE nCheck OF
                    1: bOk := bOk OR (eSt <> E_State.Aborted AND eSt <> E_State.Stopped);
                    2: bOk := bOk OR eSt = E_State.Idle;
                ELSE
                    bOk := bOk OR eSt <> E_State.Aborted;
                END_CASE
            END_IF
        END_FOR
        IF NOT bOk AND NOT (bWithdrawn AND nCheck <> 2) AND (bAny OR nCheck <> 3) THEN
            MissingGroup := g;
            RETURN;
        END_IF
    END_IF
END_FOR
END_METHOD

// Fonctions visées par une Route du process général (après chaque déploiement)
METHOD ScanGroups
VAR
    k : INT;
    g : DINT;
END_VAR
MEMSET(ADR(_aGroupUsed), 0, SIZEOF(_aGroupUsed));
FOR k := 1 TO MIN(_refMachine.nInstrCount, GVL_Const.MAX_INSTR) DO
    IF _refMachine.aInstr[k].eOp = E_Op.Route THEN
        g := _refMachine.aInstr[k].aArg[1];
        IF g >= 1 AND g <= GVL_Const.MAX_GROUPS THEN _aGroupUsed[g] := TRUE; END_IF
    END_IF
END_FOR
IF _refMachine.nRejectGroup >= 1 AND _refMachine.nRejectGroup <= GVL_Const.MAX_GROUPS THEN _aGroupUsed[_refMachine.nRejectGroup] := TRUE; END_IF
END_METHOD

// Contexte d'un mover, pour un lancement HMI d'opération avec mover (docs/05 § 8)
METHOD MoverPtr : POINTER TO ST_MoverCtx
VAR_INPUT
    nMover : USINT;
END_VAR
MoverPtr := 0;
IF nMover >= 1 AND nMover <= GVL_Const.MAX_MOVERS THEN MoverPtr := ADR(aMover[nMover]); END_IF
END_METHOD

METHOD MoverInError : BOOL
VAR
    i : USINT;
END_VAR
MoverInError := FALSE;
FOR i := 1 TO _refMachine.nMovers DO
    IF aMover[i].eState = E_MoverState.Error THEN MoverInError := TRUE; END_IF
END_FOR
END_METHOD

METHOD ClearFaults
VAR
    i : USINT;
END_VAR
bMachineFault := FALSE;
nFaultCode := 0;
FOR i := 1 TO GVL_Const.MAX_MOVERS DO
    IF aMover[i].eState = E_MoverState.Error THEN aMover[i].eState := E_MoverState.Ready; END_IF
END_FOR
END_METHOD

// Table d'OF publiée dans le statut de la machine (docs/06 § 6.3)
METHOD PublishOrders
VAR_IN_OUT
    stStatus : ST_MachineStatus;
END_VAR
stStatus.aOrder := aOrder;
stStatus.nActiveOrder := 0;
IF nActiveOrder >= 1 AND nActiveOrder <= GVL_Const.MAX_ORDERS THEN stStatus.nActiveOrder := aOrder[nActiveOrder].nOrder; END_IF
END_METHOD

METHOD PRIVATE _Publish
VAR
    i : USINT;
    k : USINT;
    stPos : ST_Position;
    ipDrv : I_PlanarDriver;
END_VAR
ipDrv := _refMgr.Driver;
FOR i := 1 TO GVL_Const.MAX_MOVERS DO
    IF ipDrv <> 0 THEN
        stPos := ipDrv.MoverPosition(i);
        aMover[i].fX := stPos.fX;
        aMover[i].fY := stPos.fY;
        aMover[i].fC := stPos.fC;
    END_IF
    GVL_Hmi.aMoverStatus[i].eState := aMover[i].eState;
    GVL_Hmi.aMoverStatus[i].eWait := aMover[i].eWait;
    GVL_Hmi.aMoverStatus[i].fX := LREAL_TO_REAL(aMover[i].fX);
    GVL_Hmi.aMoverStatus[i].fY := LREAL_TO_REAL(aMover[i].fY);
    GVL_Hmi.aMoverStatus[i].fC := LREAL_TO_REAL(aMover[i].fC);
    GVL_Hmi.aMoverStatus[i].nStation := aMover[i].nStation;
    GVL_Hmi.aMoverStatus[i].nDest := aMover[i].nDest;
    GVL_Hmi.aMoverStatus[i].nTargetGroup := aMover[i].nTargetGroup;
    GVL_Hmi.aMoverStatus[i].nTable := aMover[i].nTable;
    GVL_Hmi.aMoverStatus[i].nPC := aMover[i].nPC;
    IF aMover[i].nPC >= 1 AND aMover[i].nPC <= _refMachine.nInstrCount THEN GVL_Hmi.aMoverStatus[i].nStepId := _refMachine.aInstr[aMover[i].nPC].nStepId; END_IF
    GVL_Hmi.aMoverStatus[i].bOutOfService := aMover[i].bOutOfService;
    GVL_Hmi.aMoverStatus[i].bQualityLock := aMover[i].bQualityLock;
    GVL_Hmi.aMoverStatus[i].bAbsent := aMover[i].bAbsent;
    FOR k := 1 TO GVL_Const.MAX_SLOTS DO
        GVL_Hmi.aMoverStatus[i].aSlot[k].bPresent := aMover[i].aSlot[k].bPresent;
        GVL_Hmi.aMoverStatus[i].aSlot[k].sPartId := aMover[i].aSlot[k].sPartId;
        GVL_Hmi.aMoverStatus[i].aSlot[k].eStatus := aMover[i].aSlot[k].eStatus;
        GVL_Hmi.aMoverStatus[i].aSlot[k].eVerdict := F_Verdict(aMover[i].aSlot[k].aData[1]);
        GVL_Hmi.aMoverStatus[i].aSlot[k].nOrder := aMover[i].aSlot[k].nOrder;
    END_FOR
    GVL_Hmi.aMoverStatus[i].aVar := aMover[i].aVar;
    GVL_Hmi.aMoverStatus[i].aVarPos := aMover[i].aVarPos;
    GVL_Hmi.aMoverStatus[i].aVarId := aMover[i].aVarId;
END_FOR
END_METHOD

// ================================================================== valeurs rémanentes (docs/02 § 7.4, docs/05 § 10 étape 6)

METHOD PublishRetained
VAR_IN_OUT
    stOut : ST_RetainedValues;
END_VAR
VAR
    i : USINT;
    v : USINT;
    stItem : ST_RetainedItem;
END_VAR
FOR i := 1 TO _refMachine.nMovers DO
    FOR v := 1 TO MIN(_refMachine.nMoverVar, GVL_Const.MAX_MOVER_VARS) DO
        IF aMover[i].aVarId[v] <> 0 THEN
            MEMSET(ADR(stItem), 0, SIZEOF(stItem));
            stItem.eKind := E_RetainedKind.MoverVar;
            stItem.nMover := i;
            stItem.nId := aMover[i].aVarId[v];
            stItem.aValue[1] := aMover[i].aVar[v];
            stItem.stPos := aMover[i].aVarPos[v];
            F_AddRetained(stOut, stItem);
        END_IF
    END_FOR
END_FOR
END_METHOD

METHOD Restore : BOOL
VAR_IN_OUT
    stItem : ST_RetainedItem;
END_VAR
VAR
    v : USINT;
END_VAR
Restore := FALSE;
IF stItem.eKind <> E_RetainedKind.MoverVar OR stItem.nMover < 1 OR stItem.nMover > _refMachine.nMovers OR stItem.nId = 0 THEN RETURN; END_IF
FOR v := 1 TO MIN(_refMachine.nMoverVar, GVL_Const.MAX_MOVER_VARS) DO
    IF aMover[stItem.nMover].aVarId[v] = stItem.nId THEN
        aMover[stItem.nMover].aVar[v] := stItem.aValue[1];
        aMover[stItem.nMover].aVarPos[v] := stItem.stPos;
        Restore := TRUE;
        RETURN;
    END_IF
END_FOR
END_METHOD
END_FUNCTION_BLOCK

(* ---- FB_Loader.st ---- *)
// Chargeur (docs/05 § 10) : vérification de la zone d'attente (versions, sommes de contrôle, structure, pools),
// demande d'activation à FB_Machine, liste de restauration des valeurs rémanentes.
//
// Codes d'erreur de ST_DeployError.nCode (D94) :
//   1 jeu d'instructions demandé trop récent (nDetail = version demandée)   2 catalogue demandé trop récent
//   3 somme de contrôle fausse (nStation = bloc, 17 = recettes ; nDetail = CRC calculé)
//   4 type inconnu du catalogue du PLC (nDetail = type)   5 n° local en double, hors limites ou hors rang
//   6 parent invalide (absent ou rangé après l'enfant)   7 pool insuffisant ou type absent de la bibliothèque
//   8 signal ou élément matériel invalide (nDetail = n° de signal, 100 = élément matériel)
//   9 sortie écrite par deux objets (nDetail = index DO, 10000 + index AO)   10 instruction inconnue (nDetail = n° d'opération)
//   11 saut hors de la table   12 objet invalide   13 action invalide pour le type (nDetail = action)
//   14 condition absente   15 texte absent   16 position nommée absente   17 Fork/Join non appariés
//   18 profondeur d'appel supérieure à 4   19 table invalide (début, longueur, nature ; nDetail = table)
//   20 configuration refusée par l'objet   21 machine pas Stopped
//   22 configuration machine invalide (nDetail : 1 movers, 2 emplacements, 3 positions planaires, 4 parcage,
//      5 position d'une station, 6 fonction de rebut, 7 fonction d'une Route, 8 station d'une calibration)
FUNCTION_BLOCK FB_Loader
VAR_INPUT
    bMachineStopped : BOOL;
END_VAR
VAR_OUTPUT
    bActivate : BOOL;               // impulsion : zone d'attente vérifiée, FB_Machine l'active ce cycle puis appelle Finish
    bRestore : BOOL;                // impulsion : liste de restauration complète, FB_Machine l'applique puis appelle RestoreDone
    bBusy : BOOL;
    nRestoreCount : UINT;           // liste de restauration reçue (docs/05 § 10, étape 6)
    aRestore : ARRAY[1..2048] OF ST_RetainedItem;
    sRestoreUser : STRING(24);
END_VAR
VAR
    _refFactory : REFERENCE TO FB_ObjectFactory;
    fbCrc : FB_Crc32;
    _nLastSeq : UDINT;
    _stReq : ST_DeployRequest;
    _stResp : ST_DeployResponse;
    _nStep : USINT;                 // 0 libre, 1 sommes de contrôle, 2 structure, 3 activation demandée
    _nBlock : USINT;
    _bVerified : BOOL;
    _aDoUsed : ARRAY[0..(GVL_Const.MAX_DO / 32) - 1] OF DWORD;
    _aAoUsed : ARRAY[0..(GVL_Const.MAX_AO / 32) - 1] OF DWORD;
    // Restauration (docs/05 § 10, étape 6)
    _nLastRestoreSeq : UDINT;
    _nRestorePage : UINT;
END_VAR
VAR CONSTANT
    CRC_BUDGET : UDINT := 65536;    // octets par cycle
END_VAR

METHOD Init
VAR_INPUT
    refFactory : REFERENCE TO FB_ObjectFactory;
END_VAR
_refFactory REF= refFactory;
_nLastSeq := GVL_Hmi.stDeploy.nSeq;
_nLastRestoreSeq := GVL_Hmi.stRestore.nSeq;
END_METHOD

METHOD Cycle
VAR
    bDone : BOOL;
END_VAR
bActivate := FALSE;
bRestore := FALSE;
_Restore();

CASE _nStep OF
    0:
        IF GVL_Hmi.stDeploy.nSeq = _nLastSeq THEN RETURN; END_IF
        _nLastSeq := GVL_Hmi.stDeploy.nSeq;
        _stReq := GVL_Hmi.stDeploy;
        MEMSET(ADR(_stResp), 0, SIZEOF(_stResp));
        _stResp.nSeq := _stReq.nSeq;
        CASE _stReq.eCmd OF
            E_DeployCmd.Cancel:
                _bVerified := FALSE;
                _Respond(TRUE);
            E_DeployCmd.Verify, E_DeployCmd.Activate:
                _bVerified := FALSE;
                IF NOT bMachineStopped THEN
                    F_AddDeployError(_stResp, 21, 0, 0, 0, 0, 0);
                    _Respond(FALSE);
                    RETURN;
                END_IF
                IF _stReq.nInstrSetRequired > GVL_Const.INSTR_SET_VERSION THEN
                    F_AddDeployError(_stResp, 1, 0, 0, 0, GVL_Const.INSTR_SET_VERSION, _stReq.nInstrSetRequired);
                END_IF
                IF _stReq.nCatalogRequired > GVL_Catalog.CatalogVersion THEN
                    F_AddDeployError(_stResp, 2, 0, 0, 0, GVL_Catalog.CatalogVersion, _stReq.nCatalogRequired);
                END_IF
                IF _stResp.nErrors > 0 THEN _Respond(FALSE); RETURN; END_IF
                _nBlock := 0;
                _BeginCrc(0);
                _nStep := 1;
        ELSE
            _Respond(FALSE);
        END_CASE

    1:  // Sommes de contrôle : un bloc après l'autre, CRC_BUDGET octets par cycle
        bDone := fbCrc.Step(CRC_BUDGET);
        IF bDone THEN
            IF fbCrc.Value <> _ExpectedCrc(_nBlock) THEN F_AddDeployError(_stResp, 3, _nBlock, 0, 0, 0, fbCrc.Value); END_IF
            IF _nBlock >= GVL_Const.MAX_STATIONS + 1 THEN
                IF _stResp.nErrors > 0 THEN _Respond(FALSE); RETURN; END_IF
                MEMSET(ADR(_aDoUsed), 0, SIZEOF(_aDoUsed));
                MEMSET(ADR(_aAoUsed), 0, SIZEOF(_aAoUsed));
                _nBlock := 0;
                _nStep := 2;
            ELSE
                _nBlock := _nBlock + 1;
                _BeginCrc(_nBlock);
            END_IF
        END_IF

    2:  // Structure : un bloc par cycle, puis les pools
        IF _nBlock = 0 THEN
            _CheckMachine();
        ELSE
            _CheckStation(_nBlock);
        END_IF
        IF _nBlock < GVL_Const.MAX_STATIONS THEN
            _nBlock := _nBlock + 1;
        ELSE
            _refFactory.Check(GVL_Hmi.stStaging, _stResp);
            IF _stResp.nErrors > 0 THEN
                _Respond(FALSE);
            ELSIF _stReq.eCmd = E_DeployCmd.Verify THEN
                _bVerified := TRUE;
                _Respond(TRUE);
            ELSIF NOT bMachineStopped THEN
                F_AddDeployError(_stResp, 21, 0, 0, 0, 0, 0);
                _Respond(FALSE);
            ELSE
                bActivate := TRUE;
                _nStep := 3;
            END_IF
        END_IF

    3:  // FB_Machine active et appelle Finish
        ;
END_CASE
bBusy := _nStep <> 0;
END_METHOD

// Fin de l'activation par FB_Machine (docs/05 § 10, étapes 4 et 5)
METHOD Finish
VAR_IN_OUT
    stFactoryResp : ST_DeployResponse;
END_VAR
VAR
    k : USINT;
END_VAR
FOR k := 1 TO stFactoryResp.nErrors DO
    F_AddDeployError(_stResp, stFactoryResp.aError[k].nCode, stFactoryResp.aError[k].nStation, stFactoryResp.aError[k].nTable,
                     stFactoryResp.aError[k].nInstr, stFactoryResp.aError[k].nObject, stFactoryResp.aError[k].nDetail);
END_FOR
_Respond(_stResp.nErrors = 0);
END_METHOD

PROPERTY Request : REFERENCE TO ST_DeployRequest
GET
Request REF= _stReq;
END_GET
END_PROPERTY

METHOD PRIVATE _Respond
VAR_INPUT
    bOk : BOOL;
END_VAR
_stResp.eResult := SEL(bOk, E_CmdResult.Rejected, E_CmdResult.Accepted);
GVL_Hmi.stDeployResp := _stResp;
_nStep := 0;
bBusy := FALSE;
END_METHOD

METHOD PRIVATE _BeginCrc
VAR_INPUT
    nBlock : USINT;
END_VAR
IF nBlock = 0 THEN
    fbCrc.Begin(ADR(GVL_Hmi.stStaging.stMachine), SIZEOF(GVL_Hmi.stStaging.stMachine));
ELSIF nBlock <= GVL_Const.MAX_STATIONS THEN
    fbCrc.Begin(ADR(GVL_Hmi.stStaging.aStation[nBlock]), SIZEOF(GVL_Hmi.stStaging.aStation[nBlock]));
ELSE
    fbCrc.Begin(ADR(GVL_Hmi.stStaging.aPressRecipe), SIZEOF(GVL_Hmi.stStaging.aPressRecipe));
END_IF
END_METHOD

METHOD PRIVATE _ExpectedCrc : UDINT
VAR_INPUT
    nBlock : USINT;
END_VAR
IF nBlock = 0 THEN
    _ExpectedCrc := _stReq.nCrcMachine;
ELSIF nBlock <= GVL_Const.MAX_STATIONS THEN
    _ExpectedCrc := _stReq.aCrcStation[nBlock];
ELSE
    _ExpectedCrc := _stReq.nCrcRecipes;
END_IF
END_METHOD

// ------------------------------------------------------------------ structure

METHOD PRIVATE _CheckMachine
VAR
    m : REFERENCE TO ST_MachineData;
    s : USINT;
    q : USINT;
    k : INT;
    g : DINT;
END_VAR
m REF= GVL_Hmi.stStaging.stMachine;
IF m.nMovers > GVL_Const.MAX_MOVERS THEN F_AddDeployError(_stResp, 22, 0, 0, 0, 0, 1); END_IF
IF m.nSlots < 1 OR m.nSlots > GVL_Const.MAX_SLOTS THEN F_AddDeployError(_stResp, 22, 0, 0, 0, 0, 2); END_IF
IF m.nPlanarPos < 0 OR m.nPlanarPos > GVL_Const.MAX_PLANAR_POS THEN F_AddDeployError(_stResp, 22, 0, 0, 0, 0, 3); RETURN; END_IF
IF m.nParkPos < 0 OR m.nParkPos > m.nPlanarPos OR_ELSE (m.nParkPos > 0 AND_THEN m.aPlanarPos[m.nParkPos].eKind <> E_PlanarPosKind.Park) THEN
    F_AddDeployError(_stResp, 22, 0, 0, 0, 0, 4);
END_IF
FOR s := 1 TO GVL_Const.MAX_STATIONS DO
    IF m.aStation[s].bUsed THEN
        IF m.aStation[s].nWorkPos < 1 OR m.aStation[s].nWorkPos > m.nPlanarPos THEN F_AddDeployError(_stResp, 22, s, 0, 0, 0, 5); END_IF
        FOR q := 1 TO GVL_Const.MAX_QUEUE DO
            IF m.aStation[s].aQueuePos[q] < 0 OR m.aStation[s].aQueuePos[q] > m.nPlanarPos THEN F_AddDeployError(_stResp, 22, s, 0, 0, q, 5); END_IF
        END_FOR
    END_IF
END_FOR
IF m.nRejectGroup > GVL_Const.MAX_GROUPS OR_ELSE (m.nRejectGroup > 0 AND_THEN m.aGroup[m.nRejectGroup].eRole <> E_GroupRole.Reject) THEN
    F_AddDeployError(_stResp, 22, 0, 0, 0, 0, 6);
END_IF
FOR k := 1 TO MIN(m.nInstrCount, GVL_Const.MAX_INSTR) DO
    IF m.aInstr[k].eOp = E_Op.Route THEN
        g := m.aInstr[k].aArg[1];
        IF g < 1 OR g > GVL_Const.MAX_GROUPS OR_ELSE NOT m.aGroup[g].bUsed THEN F_AddDeployError(_stResp, 22, 0, 0, k, 0, 7); END_IF
    ELSIF m.aInstr[k].eOp = E_Op.CalibStation THEN
        g := m.aInstr[k].aArg[1];
        IF g < 1 OR g > GVL_Const.MAX_STATIONS OR_ELSE NOT m.aStation[g].bUsed THEN F_AddDeployError(_stResp, 22, 0, 0, k, 0, 8); END_IF
    END_IF
END_FOR
_CheckObjects(0, ADR(m.aMachineObj), m.nMachineObj, GVL_Const.MAX_MACHINE_OBJ);
_CheckTables(0, ADR(m.aTable), ADR(m.aInstr), m.nInstrCount, ADR(m.aCond), ADR(m.aText), ADR(m.aMachineObj), m.nMachineObj);
END_METHOD

METHOD PRIVATE _CheckStation
VAR_INPUT
    n : USINT;
END_VAR
VAR
    d : REFERENCE TO ST_StationData;
    k : USINT;
    t : USINT;
END_VAR
d REF= GVL_Hmi.stStaging.aStation[n];
IF NOT GVL_Hmi.stStaging.stMachine.aStation[n].bUsed AND d.nObjCount = 0 THEN RETURN; END_IF
_CheckObjects(n, ADR(d.aObj), d.nObjCount, GVL_Const.MAX_OBJ_PER_STATION);
_CheckTables(n, ADR(d.aTable), ADR(d.aInstr), d.nInstrCount, ADR(d.aCond), ADR(d.aText), ADR(d.aObj), d.nObjCount);
FOR k := 1 TO MIN(d.nOpMapCount, GVL_Const.MAX_OPMAP) DO
    t := d.aOpMap[k].nTable;
    IF d.aOpMap[k].nGroup < 1 OR d.aOpMap[k].nGroup > GVL_Const.MAX_GROUPS OR d.aOpMap[k].nOperationNo < 1 OR d.aOpMap[k].nOperationNo > 8
       OR t < 1 OR t > GVL_Const.MAX_TABLES OR_ELSE NOT d.aTable[t].bUsed OR_ELSE d.aTable[t].eKind <> E_TableKind.Operation THEN
        F_AddDeployError(_stResp, 19, n, t, 0, 0, k);
    END_IF
END_FOR
FOR k := 1 TO MIN(d.nCalibCount, GVL_Const.CALIB_PER_STATION) DO
    t := d.aCalib[k].nTable;
    IF t < 1 OR t > GVL_Const.MAX_TABLES OR_ELSE NOT d.aTable[t].bUsed OR_ELSE d.aTable[t].eKind <> E_TableKind.Calibration THEN
        F_AddDeployError(_stResp, 19, n, t, 0, 0, 100 + k);
    END_IF
END_FOR
END_METHOD

METHOD PRIVATE _CheckObjects
VAR_INPUT
    n : USINT;
    pObj : POINTER TO ARRAY[1..GVL_Const.MAX_OBJ_PER_STATION] OF ST_ObjConfig;
    nCount : UINT;
    nMax : UINT;
END_VAR
VAR
    k : UINT;
    s : USINT;
    o : REFERENCE TO ST_ObjConfig;
    idx : INT;
    bReal : BOOL;
END_VAR
IF nCount > nMax THEN
    F_AddDeployError(_stResp, 5, n, 0, 0, nCount, nMax);
    RETURN;
END_IF
FOR k := 1 TO nCount DO
    o REF= pObj^[k];
    // Le compilateur range les objets par n° local, parents avant enfants : rang = n° local
    IF o.nLocalId <> k THEN F_AddDeployError(_stResp, 5, n, 0, 0, k, o.nLocalId); END_IF
    IF o.nParentId >= k THEN F_AddDeployError(_stResp, 6, n, 0, 0, k, o.nParentId); END_IF
    bReal := NOT o.bSimulated AND NOT o.bDisabled;
    FOR s := 1 TO GVL_Const.MAX_SIGNALS DO
        idx := o.aSignal[s].nIndex;
        CASE o.aSignal[s].eKind OF
            E_SignalKind.DI:
                IF idx < 0 OR idx >= GVL_Const.MAX_DI THEN F_AddDeployError(_stResp, 8, n, 0, 0, k, s); END_IF
            E_SignalKind.AI:
                IF idx < 0 OR idx >= GVL_Const.MAX_AI THEN F_AddDeployError(_stResp, 8, n, 0, 0, k, s); END_IF
            E_SignalKind.DO:
                IF idx < 0 OR idx >= GVL_Const.MAX_DO THEN
                    F_AddDeployError(_stResp, 8, n, 0, 0, k, s);
                ELSIF bReal THEN
                    IF (SHR(_aDoUsed[idx / 32], idx MOD 32) AND 1) = 1 THEN F_AddDeployError(_stResp, 9, n, 0, 0, k, INT_TO_UDINT(idx)); END_IF
                    _aDoUsed[idx / 32] := _aDoUsed[idx / 32] OR SHL(DWORD#1, idx MOD 32);
                END_IF
            E_SignalKind.AO:
                IF idx < 0 OR idx >= GVL_Const.MAX_AO THEN
                    F_AddDeployError(_stResp, 8, n, 0, 0, k, s);
                ELSIF bReal THEN
                    IF (SHR(_aAoUsed[idx / 32], idx MOD 32) AND 1) = 1 THEN F_AddDeployError(_stResp, 9, n, 0, 0, k, 10000 + INT_TO_UDINT(idx)); END_IF
                    _aAoUsed[idx / 32] := _aAoUsed[idx / 32] OR SHL(DWORD#1, idx MOD 32);
                END_IF
        END_CASE
    END_FOR
    // Élément matériel : un axe réel doit désigner un axe relié dans GVL_Hw
    IF bReal AND (o.nType = GVL_Catalog.Type_LinearAxis OR o.nType = GVL_Catalog.Type_RotaryAxis)
       AND (o.nDevice < 1 OR o.nDevice > GVL_IoRef.nAxes) THEN
        F_AddDeployError(_stResp, 8, n, 0, 0, k, 100);
    END_IF
END_FOR
END_METHOD

METHOD PRIVATE _CheckTables
VAR_INPUT
    n : USINT;
    pTable : POINTER TO ARRAY[1..GVL_Const.MAX_TABLES] OF ST_TableDir;
    pInstr : POINTER TO ARRAY[1..GVL_Const.MAX_INSTR] OF ST_Instr;
    nInstrCount : INT;
    pCond : POINTER TO ARRAY[1..GVL_Const.MAX_COND] OF ST_Condition;
    pText : POINTER TO ARRAY[1..GVL_Const.MAX_TEXTS] OF STRING(80);
    pObj : POINTER TO ARRAY[1..GVL_Const.MAX_OBJ_PER_STATION] OF ST_ObjConfig;
    nObjCount : UINT;
END_VAR
VAR
    t : USINT;
    i : INT;
    nS : INT;
    nE : INT;
    p : USINT;
    b : USINT;
    ins : REFERENCE TO ST_Instr;
    nForks : INT;
    nJoins : INT;
    aDepth : ARRAY[1..GVL_Const.MAX_TABLES] OF INT;
    nPass : INT;
    nCallee : DINT;
END_VAR
IF nInstrCount < 0 OR nInstrCount > GVL_Const.MAX_INSTR THEN
    F_AddDeployError(_stResp, 19, n, 0, 0, 0, 0);
    RETURN;
END_IF
FOR t := 1 TO GVL_Const.MAX_TABLES DO
    IF pTable^[t].bUsed THEN
        nS := pTable^[t].nStart;
        nE := pTable^[t].nStart + pTable^[t].nLength - 1;
        IF nS < 1 OR pTable^[t].nLength < 1 OR nE > nInstrCount THEN
            F_AddDeployError(_stResp, 19, n, t, 0, 0, t);
        ELSE
            nForks := 0;
            nJoins := 0;
            FOR i := nS TO nE DO
                ins REF= pInstr^[i];
                IF ins.eOp > E_Op.SetOut THEN F_AddDeployError(_stResp, 10, n, t, i, 0, 0); END_IF
                CASE ins.eOp OF
                    E_Op.Jump:
                        IF NOT _In(ins.aArg[1], nS, nE) THEN F_AddDeployError(_stResp, 11, n, t, i, 0, DINT_TO_UDINT(ins.aArg[1])); END_IF
                    E_Op.JumpIfFalse:
                        IF NOT _In(ins.aArg[2], nS, nE) THEN F_AddDeployError(_stResp, 11, n, t, i, 0, DINT_TO_UDINT(ins.aArg[2])); END_IF
                        IF NOT _CondOk(pCond, ins.aArg[1]) THEN F_AddDeployError(_stResp, 14, n, t, i, 0, DINT_TO_UDINT(ins.aArg[1])); END_IF
                    E_Op.WaitCond:
                        IF NOT _CondOk(pCond, ins.aArg[1]) THEN F_AddDeployError(_stResp, 14, n, t, i, 0, DINT_TO_UDINT(ins.aArg[1])); END_IF
                    E_Op.LoopNext:
                        IF NOT _In(ins.aArg[2], nS, nE) THEN F_AddDeployError(_stResp, 11, n, t, i, 0, DINT_TO_UDINT(ins.aArg[2])); END_IF
                    E_Op.Fork:
                        nForks := nForks + 1;
                        IF NOT _In(ins.aArg[1], nS, nE) THEN
                            F_AddDeployError(_stResp, 17, n, t, i, 0, DINT_TO_UDINT(ins.aArg[1]));
                        ELSIF pInstr^[ins.aArg[1]].eOp <> E_Op.Join OR pInstr^[ins.aArg[1]].aArg[1] <> i THEN
                            F_AddDeployError(_stResp, 17, n, t, i, 0, DINT_TO_UDINT(ins.aArg[1]));
                        END_IF
                        FOR b := 2 TO 5 DO
                            IF ins.aArg[b] <> 0 AND NOT _In(ins.aArg[b], nS, nE) THEN F_AddDeployError(_stResp, 11, n, t, i, 0, DINT_TO_UDINT(ins.aArg[b])); END_IF
                        END_FOR
                    E_Op.Join:
                        nJoins := nJoins + 1;
                    E_Op.Call:
                        IF ins.aArg[1] < 1 OR ins.aArg[1] > GVL_Const.MAX_TABLES OR_ELSE NOT pTable^[ins.aArg[1]].bUsed THEN
                            F_AddDeployError(_stResp, 19, n, t, i, 0, DINT_TO_UDINT(ins.aArg[1]));
                        END_IF
                    E_Op.Action, E_Op.SavePos:
                        IF ins.nObject < 1 OR ins.nObject > nObjCount THEN
                            F_AddDeployError(_stResp, 12, n, t, i, ins.nObject, 0);
                        ELSIF ins.eOp = E_Op.Action AND_THEN NOT F_CatalogHasAction(pObj^[ins.nObject].nType, ins.nAction) THEN
                            F_AddDeployError(_stResp, 13, n, t, i, ins.nObject, ins.nAction);
                        END_IF
                    E_Op.Alarm, E_Op.Prompt:
                        IF ins.aArg[1] < 0 OR ins.aArg[1] > GVL_Const.MAX_TEXTS THEN F_AddDeployError(_stResp, 15, n, t, i, 0, DINT_TO_UDINT(ins.aArg[1])); END_IF
                END_CASE
                IF ins.eOnFail = E_FailPolicy.Goto AND NOT _In(ins.nFailTarget, nS, nE) THEN
                    F_AddDeployError(_stResp, 11, n, t, i, 0, INT_TO_UDINT(ins.nFailTarget));
                END_IF
                FOR p := 1 TO GVL_Const.MAX_PARAMS DO
                    CASE ins.aParam[p].eSource OF
                        E_ValueSource.NamedPos:
                            IF n = 0 OR ins.aParam[p].nIndex < 1 OR ins.aParam[p].nIndex > GVL_Const.MAX_NAMED_POS THEN
                                F_AddDeployError(_stResp, 16, n, t, i, 0, INT_TO_UDINT(ins.aParam[p].nIndex));
                            END_IF
                        E_ValueSource.Text:
                            IF ins.aParam[p].nIndex < 1 OR ins.aParam[p].nIndex > GVL_Const.MAX_TEXTS THEN
                                F_AddDeployError(_stResp, 15, n, t, i, 0, INT_TO_UDINT(ins.aParam[p].nIndex));
                            END_IF
                        E_ValueSource.ObjValue:
                            IF ins.aParam[p].nIndex < 1 OR ins.aParam[p].nIndex > UINT_TO_INT(nObjCount) THEN
                                F_AddDeployError(_stResp, 12, n, t, i, INT_TO_UINT(ins.aParam[p].nIndex), p);
                            END_IF
                    END_CASE
                END_FOR
            END_FOR
            IF nForks <> nJoins THEN F_AddDeployError(_stResp, 17, n, t, 0, 0, INT_TO_UDINT(nForks)); END_IF
        END_IF
    END_IF
END_FOR
// Profondeur d'appel : plus longue chaîne de Call depuis chaque table ; une boucle d'appels la fait croître sans fin
FOR nPass := 1 TO GVL_Const.MAX_CALL_DEPTH + 2 DO
    FOR t := 1 TO GVL_Const.MAX_TABLES DO
        IF pTable^[t].bUsed AND pTable^[t].nStart >= 1 THEN
            FOR i := pTable^[t].nStart TO MIN(pTable^[t].nStart + pTable^[t].nLength - 1, nInstrCount) DO
                IF pInstr^[i].eOp = E_Op.Call THEN
                    nCallee := pInstr^[i].aArg[1];
                    IF nCallee >= 1 AND nCallee <= GVL_Const.MAX_TABLES THEN aDepth[t] := MAX(aDepth[t], aDepth[nCallee] + 1); END_IF
                END_IF
            END_FOR
        END_IF
    END_FOR
END_FOR
FOR t := 1 TO GVL_Const.MAX_TABLES DO
    IF aDepth[t] > GVL_Const.MAX_CALL_DEPTH THEN F_AddDeployError(_stResp, 18, n, t, 0, 0, INT_TO_UDINT(aDepth[t])); END_IF
END_FOR
END_METHOD

METHOD PRIVATE _In : BOOL
VAR_INPUT
    nTarget : DINT;
    nS : INT;
    nE : INT;
END_VAR
_In := nTarget >= nS AND nTarget <= nE;
END_METHOD

METHOD PRIVATE _CondOk : BOOL
VAR_INPUT
    pCond : POINTER TO ARRAY[1..GVL_Const.MAX_COND] OF ST_Condition;
    n : DINT;
END_VAR
_CondOk := n >= 1 AND n <= GVL_Const.MAX_COND AND_THEN pCond^[n].nTerms >= 1 AND pCond^[n].nTerms <= GVL_Const.MAX_COND_TERMS;
END_METHOD

// ------------------------------------------------------------------ restauration (docs/05 § 10, étape 6)

METHOD PRIVATE _Restore
VAR
    req : REFERENCE TO ST_RestoreRequest;
    k : UINT;
END_VAR
req REF= GVL_Hmi.stRestore;
IF req.nSeq = _nLastRestoreSeq THEN RETURN; END_IF
_nLastRestoreSeq := req.nSeq;
GVL_Hmi.stRestoreResp.nSeq := req.nSeq;
GVL_Hmi.stRestoreResp.nDetail := 0;
IF NOT bMachineStopped OR _nStep <> 0 THEN
    GVL_Hmi.stRestoreResp.eResult := E_CmdResult.Rejected;
    GVL_Hmi.stRestoreResp.eReason := SEL(bMachineStopped, E_RejectReason.WrongState, E_RejectReason.Busy);
    RETURN;
END_IF
IF req.nPage = 0 THEN nRestoreCount := 0; END_IF
IF req.nPage <> 0 AND req.nPage <> _nRestorePage + 1 THEN
    GVL_Hmi.stRestoreResp.eResult := E_CmdResult.Rejected;      // page perdue : la HMI recommence à la page 0
    GVL_Hmi.stRestoreResp.eReason := E_RejectReason.NotAllowed;
    RETURN;
END_IF
_nRestorePage := req.nPage;
FOR k := 1 TO MIN(req.nCount, 256) DO
    IF nRestoreCount < 2048 THEN
        nRestoreCount := nRestoreCount + 1;
        aRestore[nRestoreCount] := req.aItem[k];
    END_IF
END_FOR
sRestoreUser := req.sUser;
GVL_Hmi.stRestoreResp.eResult := E_CmdResult.Accepted;
GVL_Hmi.stRestoreResp.eReason := E_RejectReason.None;
IF req.bLast THEN bRestore := TRUE; END_IF
END_METHOD

// FB_Machine a appliqué la liste : nUnknown éléments sans correspondant ont été ignorés
METHOD RestoreDone
VAR_INPUT
    nUnknown : UINT;
END_VAR
GVL_Hmi.stRestoreResp.nDetail := nUnknown;
nRestoreCount := 0;
_nRestorePage := 0;
END_METHOD
END_FUNCTION_BLOCK
